(* IEC 61131-3 sources: codesys-to-s7/tests/corpus/C2S7-TYPE-ENUM/neg, 1 file *)

(* ---- input.st ---- *)
FUNCTION_BLOCK FB_Case
VAR
    m : INT;
END_VAR
m := 1;
END_FUNCTION_BLOCK
